(* IEC 61131-3 sources: rusty/tests/lit/single/type_promotion/narrow_unsigned, 3 files *)

(* ---- difference_in_dint.st ---- *)
// RUN: %COMPILE %s && %RUN | %CHECK %s
// Narrow integer arithmetic whose result is correct in a 32-bit target.
FUNCTION main : DINT
    VAR
        a : USINT := 5;
        b : USINT := 7;
        ua : UINT := 5;
        ub : UINT := 7;
        big : USINT := 200;
        big2 : USINT := 100;
        s7 : SINT := 7;
        i : INT := 300;
        j : INT := 200;
        u2 : UDINT := 2;
        d : DINT;
        k : INT;
        l : LINT;
    END_VAR

    // Unsigned difference stored in DINT
    d := a - b;
    printf('DINT := USINT 5 - USINT 7 = %d$N', d);          // CHECK: DINT := USINT 5 - USINT 7 = -2
    d := ua - ub;
    printf('DINT := UINT 5 - UINT 7 = %d$N', d);            // CHECK-NEXT: DINT := UINT 5 - UINT 7 = -2

    // Results beyond the operand width
    d := big + big2;
    printf('USINT 200 + USINT 100 = %d$N', d);              // CHECK-NEXT: USINT 200 + USINT 100 = 300
    d := i * j;
    printf('DINT := INT 300 * INT 200 = %d$N', d);          // CHECK-NEXT: DINT := INT 300 * INT 200 = 60000
    k := i * j;
    printf('INT := INT 300 * INT 200 = %d$N', k);           // CHECK-NEXT: INT := INT 300 * INT 200 = -5536

    // A signed operand makes the operation signed
    l := a - s7;
    printf('LINT := USINT 5 - SINT 7 = %lld$N', l);         // CHECK-NEXT: LINT := USINT 5 - SINT 7 = -2

    // Two narrow unsigned operands are computed as UDINT, so a negative difference wraps in 32 bits
    printf('USINT 5 - USINT 7 < 0 = %d$N', a - b < 0);      // CHECK-NEXT: USINT 5 - USINT 7 < 0 = 0
    printf('UINT 5 - UINT 7 < 0 = %d$N', ua - ub < 0);      // CHECK-NEXT: UINT 5 - UINT 7 < 0 = 0
    l := (a - b) * 2;
    printf('LINT := (USINT 5 - USINT 7) * 2 = %lld$N', l);  // CHECK-NEXT: LINT := (USINT 5 - USINT 7) * 2 = 4294967292

    // An untyped literal next to a UDINT takes the UDINT type, so the difference wraps in 32 bits
    l := u2 - 3;
    printf('LINT := UDINT 2 - 3 = %lld$N', l);              // CHECK-NEXT: LINT := UDINT 2 - 3 = 4294967295
    l := 1 - u2;
    printf('LINT := 1 - UDINT 2 = %lld$N', l);              // CHECK-NEXT: LINT := 1 - UDINT 2 = 4294967295
    d := u2 - 3;
    printf('DINT := UDINT 2 - 3 = %d$N', d);                // CHECK-NEXT: DINT := UDINT 2 - 3 = -1
END_FUNCTION

(* ---- difference_moved_to_64_bit_or_real.st ---- *)
// RUN: %COMPILE %s && %RUN | %CHECK %s
// XFAIL: *
// Two narrow unsigned operands are computed as UDINT, so a negative difference is zero-extended into a 64-bit or real target.
FUNCTION show_lint : DINT
    VAR_INPUT
        v : LINT;
    END_VAR
    printf('LINT parameter = %lld$N', v);
END_FUNCTION

FUNCTION show_lreal : DINT
    VAR_INPUT
        v : LREAL;
    END_VAR
    printf('LREAL parameter = %f$N', v);
END_FUNCTION

FUNCTION main : DINT
    VAR
        a : USINT := 5;
        b : USINT := 7;
        ua : UINT := 5;
        ub : UINT := 7;
        lz : LINT := 0;
        l : LINT;
        r : LREAL;
        rr : REAL;
    END_VAR

    // Assignment to a 64-bit or real target
    l := a - b;
    printf('LINT := USINT 5 - USINT 7 = %lld$N', l);        // CHECK: LINT := USINT 5 - USINT 7 = -2
    l := ua - ub;
    printf('LINT := UINT 5 - UINT 7 = %lld$N', l);          // CHECK-NEXT: LINT := UINT 5 - UINT 7 = -2
    l := (a - b) * 2;
    printf('LINT := (USINT 5 - USINT 7) * 2 = %lld$N', l);  // CHECK-NEXT: LINT := (USINT 5 - USINT 7) * 2 = -4
    r := a - b;
    printf('LREAL := USINT 5 - USINT 7 = %f$N', r);         // CHECK-NEXT: LREAL := USINT 5 - USINT 7 = -2.000000
    rr := ua - ub;
    printf('REAL := UINT 5 - UINT 7 = %f$N', rr);           // CHECK-NEXT: REAL := UINT 5 - UINT 7 = -2.000000

    // Compare with a 64-bit operand
    printf('USINT 5 - USINT 7 < LINT 0 = %d$N', a - b < lz);    // CHECK-NEXT: USINT 5 - USINT 7 < LINT 0 = 1
    printf('UINT 5 - UINT 7 < LINT 0 = %d$N', ua - ub < lz);    // CHECK-NEXT: UINT 5 - UINT 7 < LINT 0 = 1

    // Argument for a 64-bit or real parameter
    show_lint(a - b);                                       // CHECK-NEXT: LINT parameter = -2
    show_lreal(ua - ub);                                    // CHECK-NEXT: LREAL parameter = -2.000000
END_FUNCTION

(* ---- product_in_udint.st ---- *)
// RUN: %COMPILE %s && %RUN | %CHECK %s
// Two narrow unsigned operands are computed as UDINT, so a product beyond the DINT range stays exact.
FUNCTION main : DINT
    VAR
        ui : UINT := 65535;
        ui2 : UINT := 65535;
        w : WORD := 16#FFFF;
        us : USINT := 255;
        r : UDINT;
        l : LINT;
    END_VAR

    r := ui * ui2;
    printf('UDINT := UINT 65535 * UINT 65535 = %u$N', r);   // CHECK: UDINT := UINT 65535 * UINT 65535 = 4294836225
    l := ui * ui2;
    printf('LINT := UINT 65535 * UINT 65535 = %lld$N', l);  // CHECK-NEXT: LINT := UINT 65535 * UINT 65535 = 4294836225
    r := ui * w;
    printf('UDINT := UINT 65535 * WORD 16#FFFF = %u$N', r); // CHECK-NEXT: UDINT := UINT 65535 * WORD 16#FFFF = 4294836225
    r := ui * us;
    printf('UDINT := UINT 65535 * USINT 255 = %u$N', r);    // CHECK-NEXT: UDINT := UINT 65535 * USINT 255 = 16711425
END_FUNCTION
